(* IEC 61131-3 sources: SafePLC-Gen-Evaluation/Evaluation Results/butane/run_05, 2 files *)

(* ---- io_declarations.st ---- *)
(* ==================================================  *)
(* PLC I/O Variable Declarations — CODESYS 3.5  *)
(* Generated by SafePLC-Gen Multimodal  *)
(* ==================================================  *)

VAR_GLOBAL
    (* --- Analog Inputs ---  *)
    TI_2909_Raw                  AT %IW0       : INT := 0;    (* TI-2909 — Temperature indicator, square box style,  *)
    TI_2917_Raw                  AT %IW2       : INT := 0;    (* TI-2917 — Temperature indicator high-high (HH flag  *)
    TT_2909_Raw                  AT %IW4       : INT := 0;    (* TT-2909 — Temperature transmitter on process inlet  *)
    TT_2911_Raw                  AT %IW6       : INT := 0;    (* TT-2911 — Temperature transmitter on outlet/right   *)
    TT_2917_Raw                  AT %IW8       : INT := 0;    (* TT-2917 — Temperature transmitter, right side top   *)
    XI_2901A_Raw                 AT %IW10      : INT := 0;    (* XI-2901A — Status indicator AVAILABLE for motor/equ  *)
    XI_2901B_Raw                 AT %IW12      : INT := 0;    (* XI-2901B — Status indicator AVAILABLE for motor/equ  *)
    (* --- Analog Outputs ---  *)
    HY_2903A_Out                 AT %QW0       : INT := 0;    (* HY-2903A — Hand relay/signal converter (circle), le  *)
    HY_2903B_Out                 AT %QW2       : INT := 0;    (* HY-2903B — Hand relay/signal converter (circle), ri  *)
    (* --- Digital Inputs ---  *)
    ESD_3200                     AT %IX0.0     : BOOL := FALSE;    (* ESD-3200 — Emergency shutdown input signal (square   *)
    HS_2901A                     AT %IX0.1     : BOOL := FALSE;    (* HS-2901A — Hand switch for motor/equipment 2901A, l  *)
    HS_2901A_ESTOP               AT %IX0.2     : BOOL := FALSE;    (* HS-2901A-ESTOP — Hand switch EMERGENCY STOP (circle symbo  *)
    HS_2901A_START               AT %IX0.3     : BOOL := FALSE;    (* HS-2901A-START — Hand switch START/STOP (circle symbol, f  *)
    HS_2901A1                    AT %IX0.4     : BOOL := FALSE;    (* HS-2901A1 — Hand switch LOCAL/REMOTE selector for mo  *)
    HS_2901A2                    AT %IX0.5     : BOOL := FALSE;    (* HS-2901A2 — Hand switch STOP/START for motor 2901A,   *)
    HS_2901B                     AT %IX0.6     : BOOL := FALSE;    (* HS-2901B — Hand switch for motor/equipment 2901B, r  *)
    HS_2901B_ESTOP               AT %IX0.7     : BOOL := FALSE;    (* HS-2901B-ESTOP — Hand switch EMERGENCY STOP (circle symbo  *)
    HS_2901B_START               AT %IX1.0     : BOOL := FALSE;    (* HS-2901B-START — Hand switch START/STOP (circle symbol, f  *)
    HS_2901B1                    AT %IX1.1     : BOOL := FALSE;    (* HS-2901B1 — Hand switch LOCAL/REMOTE selector for mo  *)
    HS_2901B2                    AT %IX1.2     : BOOL := FALSE;    (* HS-2901B2 — Hand switch STOP/START for motor 2901B,   *)
    PSD_2917                     AT %IX1.3     : BOOL := FALSE;    (* PSD-2917 — Pressure shutdown switch/device, square   *)
    VSHH_2901A                   AT %IX1.4     : BOOL := FALSE;    (* VSHH-2901A — Vibration switch high-high on pump/motor  *)
    VSHH_2901B                   AT %IX1.5     : BOOL := FALSE;    (* VSHH-2901B — Vibration switch high-high on pump/motor  *)
    (* --- Digital Outputs ---  *)
    KV_2904                      AT %QX0.0     : BOOL := FALSE;    (* KV-2904 — Time/schedule-controlled valve or soleno  *)
END_VAR

(* ---- generated_code.st ---- *)
(* Generated by SafePLC-Gen Multimodal — CODESYS 3.5 *)
(* IEC 61131-3 Structured Text *)
(* Date: 2026-04-25T12:21:09.815350 *)

PROGRAM MotorCoolingControl

VAR
    TI_2909_Raw                  AT %IW0       : INT := 0;
    TI_2917_Raw                  AT %IW2       : INT := 0;
    TT_2909_Raw                  AT %IW4       : INT := 0;
    TT_2911_Raw                  AT %IW6       : INT := 0;
    TT_2917_Raw                  AT %IW8       : INT := 0;
    XI_2901A_Raw                 AT %IW10      : INT := 0;
    XI_2901B_Raw                 AT %IW12      : INT := 0;
    HY_2903A_Out                 AT %QW0       : INT := 0;
    HY_2903B_Out                 AT %QW2       : INT := 0;
    ESD_3200                     AT %IX0.0     : BOOL := FALSE;
    HS_2901A                     AT %IX0.1     : BOOL := FALSE;
    HS_2901A_ESTOP               AT %IX0.2     : BOOL := FALSE;
    HS_2901A_START               AT %IX0.3     : BOOL := FALSE;
    HS_2901A1                    AT %IX0.4     : BOOL := FALSE;
    HS_2901A2                    AT %IX0.5     : BOOL := FALSE;
    HS_2901B                     AT %IX0.6     : BOOL := FALSE;
    HS_2901B_ESTOP               AT %IX0.7     : BOOL := FALSE;
    HS_2901B_START               AT %IX1.0     : BOOL := FALSE;
    HS_2901B1                    AT %IX1.1     : BOOL := FALSE;
    HS_2901B2                    AT %IX1.2     : BOOL := FALSE;
    PSD_2917                     AT %IX1.3     : BOOL := FALSE;
    VSHH_2901A                   AT %IX1.4     : BOOL := FALSE;
    VSHH_2901B                   AT %IX1.5     : BOOL := FALSE;
    KV_2904                      AT %QX0.0     : BOOL := FALSE;
END_VAR

VAR
    ESTOP                        : BOOL := FALSE;
    MANUAL_RESET                 : BOOL := FALSE;
    LOOP_2917_SAFETY_TRIP        : BOOL := TRUE;
    LOOP_2901A_TRIP              : BOOL := TRUE;
    LOOP_2901B_TRIP              : BOOL := TRUE;
    LOOP_3200_TRIP               : BOOL := TRUE;
    TT_2917_HH                   : BOOL := FALSE;
    TT_2917_LL                   : BOOL := FALSE;
    VSHH_2901A_HH                : BOOL := FALSE;
    VSHH_2901A_LL                : BOOL := FALSE;
    VSHH_2901B_HH                : BOOL := FALSE;
    VSHH_2901B_LL                : BOOL := FALSE;
    ESD_3200_HH                  : BOOL := FALSE;
    ESD_3200_LL                  : BOOL := FALSE;
    SAFE_STATE                   : BOOL := TRUE;
    FirstScan                    : BOOL := TRUE;

    Motor_2901A_Out              : BOOL := FALSE;
    Motor_2901B_Out              : BOOL := FALSE;
    MCC_Trip_Out                 : BOOL := FALSE;
    PSD_Trip_Out                 : BOOL := FALSE;

    TI_2909_Scaled               : REAL := 0.0;
    TI_2917_Scaled               : REAL := 0.0;
    TT_2909_Scaled               : REAL := 0.0;
    TT_2911_Scaled               : REAL := 0.0;
    TT_2917_Scaled               : REAL := 0.0;
    XI_2901A_Scaled              : REAL := 0.0;
    XI_2901B_Scaled              : REAL := 0.0;

    TI_2909_HH_SP                : REAL := 90.0;
    TI_2909_H_SP                 : REAL := 80.0;
    TI_2909_L_SP                 : REAL := 10.0;
    TI_2909_LL_SP                : REAL := 5.0;
    TI_2909_Deadband             : REAL := 2.0;
    TI_2909_H                    : BOOL := FALSE;
    TI_2909_L                    : BOOL := FALSE;
    TI_2909_HH_Latch             : SR := (S1 := FALSE, R := FALSE);
    TI_2909_LL_Latch             : SR := (S1 := FALSE, R := FALSE);
    TI_2909_HH_Ack               : BOOL := FALSE;
    TI_2909_LL_Ack               : BOOL := FALSE;

    TT_2909_HH_SP                : REAL := 90.0;
    TT_2909_H_SP                 : REAL := 80.0;
    TT_2909_L_SP                 : REAL := 10.0;
    TT_2909_LL_SP                : REAL := 5.0;
    TT_2909_Deadband             : REAL := 2.0;
    TT_2909_H                    : BOOL := FALSE;
    TT_2909_L                    : BOOL := FALSE;
    TT_2909_HH_Latch             : SR := (S1 := FALSE, R := FALSE);
    TT_2909_LL_Latch             : SR := (S1 := FALSE, R := FALSE);
    TT_2909_HH_Ack               : BOOL := FALSE;
    TT_2909_LL_Ack               : BOOL := FALSE;

    TT_2911_HH_SP                : REAL := 90.0;
    TT_2911_H_SP                 : REAL := 80.0;
    TT_2911_L_SP                 : REAL := 10.0;
    TT_2911_LL_SP                : REAL := 5.0;
    TT_2911_Deadband             : REAL := 2.0;
    TT_2911_H                    : BOOL := FALSE;
    TT_2911_L                    : BOOL := FALSE;
    TT_2911_HH_Latch             : SR := (S1 := FALSE, R := FALSE);
    TT_2911_LL_Latch             : SR := (S1 := FALSE, R := FALSE);
    TT_2911_HH_Ack               : BOOL := FALSE;
    TT_2911_LL_Ack               : BOOL := FALSE;

    TT_2917_HH_SP                : REAL := 95.0;
    TT_2917_H_SP                 : REAL := 85.0;
    TT_2917_L_SP                 : REAL := 10.0;
    TT_2917_LL_SP                : REAL := 5.0;
    TT_2917_Deadband             : REAL := 2.0;
    TT_2917_H                    : BOOL := FALSE;
    TT_2917_L                    : BOOL := FALSE;
    TT_2917_HH_Latch             : SR := (S1 := FALSE, R := FALSE);
    TT_2917_LL_Latch             : SR := (S1 := FALSE, R := FALSE);
    TT_2917_HH_Ack               : BOOL := FALSE;
    TT_2917_LL_Ack               : BOOL := FALSE;

    TI_2917_HH_SP                : REAL := 95.0;
    TI_2917_H_SP                 : REAL := 85.0;
    TI_2917_L_SP                 : REAL := 10.0;
    TI_2917_LL_SP                : REAL := 5.0;
    TI_2917_Deadband             : REAL := 2.0;
    TI_2917_H                    : BOOL := FALSE;
    TI_2917_L                    : BOOL := FALSE;
    TI_2917_HH_Latch             : SR := (S1 := FALSE, R := FALSE);
    TI_2917_LL_Latch             : SR := (S1 := FALSE, R := FALSE);
    TI_2917_HH_Ack               : BOOL := FALSE;
    TI_2917_LL_Ack               : BOOL := FALSE;

    XI_2901A_HH_SP               : REAL := 90.0;
    XI_2901A_H_SP                : REAL := 80.0;
    XI_2901A_L_SP                : REAL := 20.0;
    XI_2901A_LL_SP               : REAL := 10.0;
    XI_2901A_Deadband            : REAL := 2.0;
    XI_2901A_H                   : BOOL := FALSE;
    XI_2901A_L                   : BOOL := FALSE;
    XI_2901A_HH_Latch            : SR := (S1 := FALSE, R := FALSE);
    XI_2901A_LL_Latch            : SR := (S1 := FALSE, R := FALSE);
    XI_2901A_HH_Ack              : BOOL := FALSE;
    XI_2901A_LL_Ack              : BOOL := FALSE;

    XI_2901B_HH_SP               : REAL := 90.0;
    XI_2901B_H_SP                : REAL := 80.0;
    XI_2901B_L_SP                : REAL := 20.0;
    XI_2901B_LL_SP               : REAL := 10.0;
    XI_2901B_Deadband            : REAL := 2.0;
    XI_2901B_H                   : BOOL := FALSE;
    XI_2901B_L                   : BOOL := FALSE;
    XI_2901B_HH_Latch            : SR := (S1 := FALSE, R := FALSE);
    XI_2901B_LL_Latch            : SR := (S1 := FALSE, R := FALSE);
    XI_2901B_HH_Ack              : BOOL := FALSE;
    XI_2901B_LL_Ack              : BOOL := FALSE;

    HY_2903A_SP                  : REAL := 60.0;
    HY_2903A_Kp                  : REAL := 1.5;
    HY_2903A_Ki                  : REAL := 0.05;
    HY_2903A_Integral            : REAL := 0.0;
    HY_2903A_Error               : REAL := 0.0;
    HY_2903A_Output              : REAL := 0.0;

    HY_2903B_SP                  : REAL := 60.0;
    HY_2903B_Kp                  : REAL := 1.5;
    HY_2903B_Ki                  : REAL := 0.05;
    HY_2903B_Integral            : REAL := 0.0;
    HY_2903B_Error               : REAL := 0.0;
    HY_2903B_Output              : REAL := 0.0;

    Motor_2901A_Run              : BOOL := FALSE;
    Motor_2901B_Run              : BOOL := FALSE;
    Motor_2901A_StartEdge        : R_TRIG := (CLK := FALSE);
    Motor_2901B_StartEdge        : R_TRIG := (CLK := FALSE);
    Motor_2901A_StopEdge         : R_TRIG := (CLK := FALSE);
    Motor_2901B_StopEdge         : R_TRIG := (CLK := FALSE);
    Motor_2901A_StartDelay       : TON := (IN := FALSE, PT := T#3S);
    Motor_2901B_StartDelay       : TON := (IN := FALSE, PT := T#3S);
    Motor_2901A_StopCmd          : BOOL := FALSE;
    Motor_2901B_StopCmd          : BOOL := FALSE;

    System_Alarm                 : BOOL := FALSE;
END_VAR

IF FirstScan THEN
    LOOP_2917_SAFETY_TRIP := TRUE;
    LOOP_2901A_TRIP       := TRUE;
    LOOP_2901B_TRIP       := TRUE;
    LOOP_3200_TRIP        := TRUE;
    SAFE_STATE            := TRUE;
    HY_2903A_Out          := 6554;
    HY_2903B_Out          := 6554;
    KV_2904               := FALSE;
    Motor_2901A_Out       := FALSE;
    Motor_2901B_Out       := FALSE;
    MCC_Trip_Out          := TRUE;
    PSD_Trip_Out          := FALSE;
    FirstScan             := FALSE;
    RETURN;
END_IF;

ESTOP := HS_2901A_ESTOP OR HS_2901B_ESTOP OR ESD_3200;

TI_2909_Scaled  := ((INT_TO_REAL(TI_2909_Raw)  - 6554.0) / (32767.0 - 6554.0)) * 150.0;
TI_2917_Scaled  := ((INT_TO_REAL(TI_2917_Raw)  - 6554.0) / (32767.0 - 6554.0)) * 150.0;
TT_2909_Scaled  := ((INT_TO_REAL(TT_2909_Raw)  - 6554.0) / (32767.0 - 6554.0)) * 150.0;
TT_2911_Scaled  := ((INT_TO_REAL(TT_2911_Raw)  - 6554.0) / (32767.0 - 6554.0)) * 150.0;
TT_2917_Scaled  := ((INT_TO_REAL(TT_2917_Raw)  - 6554.0) / (32767.0 - 6554.0)) * 150.0;
XI_2901A_Scaled := ((INT_TO_REAL(XI_2901A_Raw) - 6554.0) / (32767.0 - 6554.0)) * 100.0;
XI_2901B_Scaled := ((INT_TO_REAL(XI_2901B_Raw) - 6554.0) / (32767.0 - 6554.0)) * 100.0;

TT_2917_HH := (TT_2917_Scaled > TT_2917_HH_SP) OR PSD_2917;
TT_2917_LL := TT_2917_Scaled < TT_2917_LL_SP;

VSHH_2901A_HH := VSHH_2901A;
VSHH_2901A_LL := FALSE;

VSHH_2901B_HH := VSHH_2901B;
VSHH_2901B_LL := FALSE;

ESD_3200_HH := ESD_3200;
ESD_3200_LL := FALSE;

IF TT_2917_HH OR TT_2917_LL THEN
    LOOP_2917_SAFETY_TRIP := TRUE;
ELSIF LOOP_2917_SAFETY_TRIP AND MANUAL_RESET
      AND NOT TT_2917_HH AND NOT TT_2917_LL THEN
    LOOP_2917_SAFETY_TRIP := FALSE;
END_IF;

IF VSHH_2901A_HH OR VSHH_2901A_LL THEN
    LOOP_2901A_TRIP := TRUE;
ELSIF LOOP_2901A_TRIP AND MANUAL_RESET
      AND NOT VSHH_2901A_HH AND NOT VSHH_2901A_LL THEN
    LOOP_2901A_TRIP := FALSE;
END_IF;

IF VSHH_2901B_HH OR VSHH_2901B_LL THEN
    LOOP_2901B_TRIP := TRUE;
ELSIF LOOP_2901B_TRIP AND MANUAL_RESET
      AND NOT VSHH_2901B_HH AND NOT VSHH_2901B_LL THEN
    LOOP_2901B_TRIP := FALSE;
END_IF;

IF ESD_3200_HH OR ESD_3200_LL THEN
    LOOP_3200_TRIP := TRUE;
ELSIF LOOP_3200_TRIP AND MANUAL_RESET
      AND NOT ESD_3200_HH AND NOT ESD_3200_LL THEN
    LOOP_3200_TRIP := FALSE;
END_IF;

SAFE_STATE := ESTOP
              OR LOOP_2917_SAFETY_TRIP
              OR LOOP_2901A_TRIP
              OR LOOP_2901B_TRIP
              OR LOOP_3200_TRIP;

IF TI_2909_Scaled >= TI_2909_HH_SP THEN
    TI_2909_HH_Latch.S1 := TRUE;
ELSIF TI_2909_Scaled <= (TI_2909_HH_SP - TI_2909_Deadband) THEN
    TI_2909_HH_Latch.S1 := FALSE;
END_IF;
TI_2909_HH_Latch.R := TI_2909_HH_Ack AND (TI_2909_Scaled < TI_2909_HH_SP);
TI_2909_HH_Latch(S1 := TI_2909_HH_Latch.S1, R := TI_2909_HH_Latch.R);
TI_2909_H := TI_2909_Scaled >= TI_2909_H_SP;
TI_2909_L := TI_2909_Scaled <= TI_2909_L_SP;
IF TI_2909_Scaled <= TI_2909_LL_SP THEN
    TI_2909_LL_Latch.S1 := TRUE;
ELSIF TI_2909_Scaled >= (TI_2909_LL_SP + TI_2909_Deadband) THEN
    TI_2909_LL_Latch.S1 := FALSE;
END_IF;
TI_2909_LL_Latch.R := TI_2909_LL_Ack AND (TI_2909_Scaled > TI_2909_LL_SP);
TI_2909_LL_Latch(S1 := TI_2909_LL_Latch.S1, R := TI_2909_LL_Latch.R);

IF TT_2909_Scaled >= TT_2909_HH_SP THEN
    TT_2909_HH_Latch.S1 := TRUE;
ELSIF TT_2909_Scaled <= (TT_2909_HH_SP - TT_2909_Deadband) THEN
    TT_2909_HH_Latch.S1 := FALSE;
END_IF;
TT_2909_HH_Latch.R := TT_2909_HH_Ack AND (TT_2909_Scaled < TT_2909_HH_SP);
TT_2909_HH_Latch(S1 := TT_2909_HH_Latch.S1, R := TT_2909_HH_Latch.R);
TT_2909_H := TT_2909_Scaled >= TT_2909_H_SP;
TT_2909_L := TT_2909_Scaled <= TT_2909_L_SP;
IF TT_2909_Scaled <= TT_2909_LL_SP THEN
    TT_2909_LL_Latch.S1 := TRUE;
ELSIF TT_2909_Scaled >= (TT_2909_LL_SP + TT_2909_Deadband) THEN
    TT_2909_LL_Latch.S1 := FALSE;
END_IF;
TT_2909_LL_Latch.R := TT_2909_LL_Ack AND (TT_2909_Scaled > TT_2909_LL_SP);
TT_2909_LL_Latch(S1 := TT_2909_LL_Latch.S1, R := TT_2909_LL_Latch.R);

IF TT_2911_Scaled >= TT_2911_HH_SP THEN
    TT_2911_HH_Latch.S1 := TRUE;
ELSIF TT_2911_Scaled <= (TT_2911_HH_SP - TT_2911_Deadband) THEN
    TT_2911_HH_Latch.S1 := FALSE;
END_IF;
TT_2911_HH_Latch.R := TT_2911_HH_Ack AND (TT_2911_Scaled < TT_2911_HH_SP);
TT_2911_HH_Latch(S1 := TT_2911_HH_Latch.S1, R := TT_2911_HH_Latch.R);
TT_2911_H := TT_2911_Scaled >= TT_2911_H_SP;
TT_2911_L := TT_2911_Scaled <= TT_2911_L_SP;
IF TT_2911_Scaled <= TT_2911_LL_SP THEN
    TT_2911_LL_Latch.S1 := TRUE;
ELSIF TT_2911_Scaled >= (TT_2911_LL_SP + TT_2911_Deadband) THEN
    TT_2911_LL_Latch.S1 := FALSE;
END_IF;
TT_2911_LL_Latch.R := TT_2911_LL_Ack AND (TT_2911_Scaled > TT_2911_LL_SP);
TT_2911_LL_Latch(S1 := TT_2911_LL_Latch.S1, R := TT_2911_LL_Latch.R);

IF TT_2917_Scaled >= TT_2917_HH_SP THEN
    TT_2917_HH_Latch.S1 := TRUE;
ELSIF TT_2917_Scaled <= (TT_2917_HH_SP - TT_2917_Deadband) THEN
    TT_2917_HH_Latch.S1 := FALSE;
END_IF;
TT_2917_HH_Latch.R := TT_2917_HH_Ack AND (TT_2917_Scaled < TT_2917_HH_SP);
TT_2917_HH_Latch(S1 := TT_2917_HH_Latch.S1, R := TT_2917_HH_Latch.R);
TT_2917_H := TT_2917_Scaled >= TT_2917_H_SP;
TT_2917_L := TT_2917_Scaled <= TT_2917_L_SP;
IF TT_2917_Scaled <= TT_2917_LL_SP THEN
    TT_2917_LL_Latch.S1 := TRUE;
ELSIF TT_2917_Scaled >= (TT_2917_LL_SP + TT_2917_Deadband) THEN
    TT_2917_LL_Latch.S1 := FALSE;
END_IF;
TT_2917_LL_Latch.R := TT_2917_LL_Ack AND (TT_2917_Scaled > TT_2917_LL_SP);
TT_2917_LL_Latch(S1 := TT_2917_LL_Latch.S1, R := TT_2917_LL_Latch.R);

IF TI_2917_Scaled >= TI_2917_HH_SP THEN
    TI_2917_HH_Latch.S1 := TRUE;
ELSIF TI_2917_Scaled <= (TI_2917_HH_SP - TI_2917_Deadband) THEN
    TI_2917_HH_Latch.S1 := FALSE;
END_IF;
TI_2917_HH_Latch.R := TI_2917_HH_Ack AND (TI_2917_Scaled < TI_2917_HH_SP);
TI_2917_HH_Latch(S1 := TI_2917_HH_Latch.S1, R := TI_2917_HH_Latch.R);
TI_2917_H := TI_2917_Scaled >= TI_2917_H_SP;
TI_2917_L := TI_2917_Scaled <= TI_2917_L_SP;
IF TI_2917_Scaled <= TI_2917_LL_SP THEN
    TI_2917_LL_Latch.S1 := TRUE;
ELSIF TI_2917_Scaled >= (TI_2917_LL_SP + TI_2917_Deadband) THEN
    TI_2917_LL_Latch.S1 := FALSE;
END_IF;
TI_2917_LL_Latch.R := TI_2917_LL_Ack AND (TI_2917_Scaled > TI_2917_LL_SP);
TI_2917_LL_Latch(S1 := TI_2917_LL_Latch.S1, R := TI_2917_LL_Latch.R);

IF XI_2901A_Scaled >= XI_2901A_HH_SP THEN
    XI_2901A_HH_Latch.S1 := TRUE;
ELSIF XI_2901A_Scaled <= (XI_2901A_HH_SP - XI_2901A_Deadband) THEN
    XI_2901A_HH_Latch.S1 := FALSE;
END_IF;
XI_2901A_HH_Latch.R := XI_2901A_HH_Ack AND (XI_2901A_Scaled < XI_2901A_HH_SP);
XI_2901A_HH_Latch(S1 := XI_2901A_HH_Latch.S1, R := XI_2901A_HH_Latch.R);
XI_2901A_H := XI_2901A_Scaled >= XI_2901A_H_SP;
XI_2901A_L := XI_2901A_Scaled <= XI_2901A_L_SP;
IF XI_2901A_Scaled <= XI_2901A_LL_SP THEN
    XI_2901A_LL_Latch.S1 := TRUE;
ELSIF XI_2901A_Scaled >= (XI_2901A_LL_SP + XI_2901A_Deadband) THEN
    XI_2901A_LL_Latch.S1 := FALSE;
END_IF;
XI_2901A_LL_Latch.R := XI_2901A_LL_Ack AND (XI_2901A_Scaled > XI_2901A_LL_SP);
XI_2901A_LL_Latch(S1 := XI_2901A_LL_Latch.S1, R := XI_2901A_LL_Latch.R);

IF XI_2901B_Scaled >= XI_2901B_HH_SP THEN
    XI_2901B_HH_Latch.S1 := TRUE;
ELSIF XI_2901B_Scaled <= (XI_2901B_HH_SP - XI_2901B_Deadband) THEN
    XI_2901B_HH_Latch.S1 := FALSE;
END_IF;
XI_2901B_HH_Latch.R := XI_2901B_HH_Ack AND (XI_2901B_Scaled < XI_2901B_HH_SP);
XI_2901B_HH_Latch(S1 := XI_2901B_HH_Latch.S1, R := XI_2901B_HH_Latch.R);
XI_2901B_H := XI_2901B_Scaled >= XI_2901B_H_SP;
XI_2901B_L := XI_2901B_Scaled <= XI_2901B_L_SP;
IF XI_2901B_Scaled <= XI_2901B_LL_SP THEN
    XI_2901B_LL_Latch.S1 := TRUE;
ELSIF XI_2901B_Scaled >= (XI_2901B_LL_SP + XI_2901B_Deadband) THEN
    XI_2901B_LL_Latch.S1 := FALSE;
END_IF;
XI_2901B_LL_Latch.R := XI_2901B_LL_Ack AND (XI_2901B_Scaled > XI_2901B_LL_SP);
XI_2901B_LL_Latch(S1 := XI_2901B_LL_Latch.S1, R := XI_2901B_LL_Latch.R);

Motor_2901A_StartEdge(CLK := HS_2901A_START OR HS_2901A OR HS_2901A2);
Motor_2901A_StopEdge(CLK  := HS_2901A_ESTOP OR HS_2901A1);
Motor_2901A_StopCmd := HS_2901A_ESTOP OR HS_2901A1;

IF Motor_2901A_StartEdge.Q AND NOT Motor_2901A_StopCmd AND NOT SAFE_STATE THEN
    Motor_2901A_Run := TRUE;
END_IF;
IF Motor_2901A_StopEdge.Q OR SAFE_STATE THEN
    Motor_2901A_Run := FALSE;
END_IF;

Motor_2901A_StartDelay(IN := Motor_2901A_Run AND NOT SAFE_STATE, PT := T#3S);

Motor_2901B_StartEdge(CLK := HS_2901B_START OR HS_2901B OR HS_2901B2);
Motor_2901B_StopEdge(CLK  := HS_2901B_ESTOP OR HS_2901B1);
Motor_2901B_StopCmd := HS_2901B_ESTOP OR HS_2901B1;

IF Motor_2901B_StartEdge.Q AND NOT Motor_2901B_StopCmd AND NOT SAFE_STATE THEN
    Motor_2901B_Run := TRUE;
END_IF;
IF Motor_2901B_StopEdge.Q OR SAFE_STATE THEN
    Motor_2901B_Run := FALSE;
END_IF;

Motor_2901B_StartDelay(IN := Motor_2901B_Run AND NOT SAFE_STATE, PT := T#3S);

IF NOT SAFE_STATE THEN
    Motor_2901A_Out  := Motor_2901A_StartDelay.Q;
    Motor_2901B_Out  := Motor_2901B_StartDelay.Q;
    MCC_Trip_Out     := FALSE;
    PSD_Trip_Out     := NOT (TT_2917_HH_Latch.Q1 OR TI_2917_HH_Latch.Q1 OR PSD_2917);
    KV_2904          := Motor_2901A_Out OR Motor_2901B_Out;

    HY_2903A_Error    := HY_2903A_SP - TT_2911_Scaled;
    HY_2903A_Integral := HY_2903A_Integral + (HY_2903A_Ki * HY_2903A_Error);
    IF HY_2903A_Integral > 100.0 THEN
        HY_2903A_Integral := 100.0;
    ELSIF HY_2903A_Integral < 0.0 THEN
        HY_2903A_Integral := 0.0;
    END_IF;
    HY_2903A_Output := (HY_2903A_Kp * HY_2903A_Error) + HY_2903A_Integral;
    IF HY_2903A_Output > 100.0 THEN
        HY_2903A_Output := 100.0;
    ELSIF HY_2903A_Output < 0.0 THEN
        HY_2903A_Output := 0.0;
    END_IF;
    HY_2903A_Out := REAL_TO_INT(6554.0 + (HY_2903A_Output / 100.0) * (32767.0 - 6554.0));

    HY_2903B_Error    := HY_2903B_SP - TT_2909_Scaled;
    HY_2903B_Integral := HY_2903B_Integral + (HY_2903B_Ki * HY_2903B_Error);
    IF HY_2903B_Integral > 100.0 THEN
        HY_2903B_Integral := 100.0;
    ELSIF HY_2903B_Integral < 0.0 THEN
        HY_2903B_Integral := 0.0;
    END_IF;
    HY_2903B_Output := (HY_2903B_Kp * HY_2903B_Error) + HY_2903B_Integral;
    IF HY_2903B_Output > 100.0 THEN
        HY_2903B_Output := 100.0;
    ELSIF HY_2903B_Output < 0.0 THEN
        HY_2903B_Output := 0.0;
    END_IF;
    HY_2903B_Out := REAL_TO_INT(6554.0 + (HY_2903B_Output / 100.0) * (32767.0 - 6554.0));
ELSE
    HY_2903A_Out      := 6554;
    HY_2903B_Out      := 6554;
    KV_2904           := FALSE;
    Motor_2901A_Out   := FALSE;
    Motor_2901B_Out   := FALSE;
    MCC_Trip_Out      := TRUE;
    PSD_Trip_Out      := FALSE;
    HY_2903A_Integral := 0.0;
    HY_2903B_Integral := 0.0;
END_IF;

System_Alarm :=
    TI_2909_HH_Latch.Q1  OR TI_2909_LL_Latch.Q1  OR TI_2909_H  OR TI_2909_L  OR
    TT_2909_HH_Latch.Q1  OR TT_2909_LL_Latch.Q1  OR TT_2909_H  OR TT_2909_L  OR
    TT_2911_HH_Latch.Q1  OR TT_2911_LL_Latch.Q1  OR TT_2911_H  OR TT_2911_L  OR
    TT_2917_HH_Latch.Q1  OR TT_2917_LL_Latch.Q1  OR TT_2917_H  OR TT_2917_L  OR
    TI_2917_HH_Latch.Q1  OR TI_2917_LL_Latch.Q1  OR TI_2917_H  OR TI_2917_L  OR
    XI_2901A_HH_Latch.Q1 OR XI_2901A_LL_Latch.Q1 OR XI_2901A_H OR XI_2901A_L OR
    XI_2901B_HH_Latch.Q1 OR XI_2901B_LL_Latch.Q1 OR XI_2901B_H OR XI_2901B_L OR
    SAFE_STATE OR MCC_Trip_Out OR PSD_Trip_Out OR Motor_2901A_Out OR Motor_2901B_Out;

END_PROGRAM
